FUNCTION_BLOCK AIWS_TO_AIS (* Composite FB for converting AIWS (WSTRING) adapter to AIS (STRING) adapter *)
  (* Standard: 61499-2; Description: Copyright (c) 2026 HR Agrartechnik GmbH This program and the accompanying materials are made available under the terms of the Eclipse Public License 2.0 which is available at https://www.eclipse.org/legal/epl-2.0/ SPDX-License-Identifier: EPL-2.0 *)
  (* Version 1.0, 2026-11-13, Franz Höpfinger, HR Agrartechnik GmbH, Initial Version - Luecke in der Adapter-Familie geschlossen *)
  PACKAGE adapter::conversion::unidirectional;
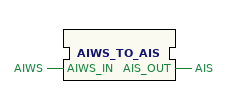
  SOCKETS
    AIWS_IN : adapter::types::unidirectional::AIWS; (* WSTRING Adapter Input *)
  END_SOCKETS
  PLUGS
    AIS_OUT : adapter::types::unidirectional::AIS; (* STRING Adapter Output *)
  END_PLUGS
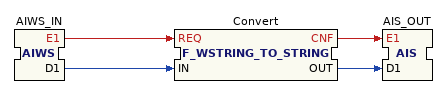
  FBS
    Convert : iec61131::conversion::F_WSTRING_TO_STRING;
  END_FBS
  EVENT_CONNECTIONS
    AIWS_IN.E1 TO Convert.REQ;
    Convert.CNF TO AIS_OUT.E1;
  END_CONNECTIONS
  DATA_CONNECTIONS
    AIWS_IN.D1 TO Convert.IN;
    Convert.OUT TO AIS_OUT.D1;
  END_CONNECTIONS
END_FUNCTION_BLOCK
